Fanuc KAREL source: KT00834.KL

PROGRAM KT00834
%NOLOCKGROUP
VAR
  R1: REAL
  R2: REAL
  OUT: INTEGER
BEGIN
  R1 = 2.0
  R2 = 3.0
  R1 = 2.0
  R2 = 3.0
  OUT = SQRT(R1)
END KT00834
